Staubli VAL3: HMI_util.dtx

mdesc mNomSpeed
public string sShowType[6]
public string sShowNum[6]
public string sJoint[6]
  [0] = "J1:"
  [1] = "J2:"
  [2] = "J3:"
  [3] = "J4:"
  [4] = "J5:"
  [5] = "J6:"
public string sCartisiam[6]
  [0] = "X:"
  [1] = "Y:"
  [2] = "Z:"
  [3] = "RX:"
  [4] = "RY:"
  [5] = "RZ:"
public string sPage
string sInputPswd
bool bConfirm
bool bCancel
string sPassword = "1"
num nUsingTool
